(* Logix 5000 project; controller TFF vendor 1 type 14 code 107 rev 34.11; software revision 34.03; part 35 of 36 *)
(* tags used below, declared in another part *)
   Config : Configuration;   // Index Array used in configuration routines
   Index : DINT;   // Index
   FirstScanComplete : BOOL;   // First Scan Complete Flag
   FlowPath : FlowPath[64];   // Flow Path Array
   FlowPathControl : FlowPathControl;   // Flow Path Control
   FlowPathSetup : FlowPathSetup;   // Flow Path Setup Data
   LI001 : ALIAS FOR AnalogPoint[44];   // Feed Bag Volume
   LI001Alarm : ALIAS FOR AlarmAnalog[44];   // Feed Bag Volume Alarm
   Phase0 : ALIAS FOR Phase[0];   // Phase 0
   SysControl : SysControl;   // General system status and command
   Tank : TankManagement;   // Tank Management
   Valve : Valve[100];   // Valve Array
   ValveControl : ValveControl;   // Valve Control
   WI001 : ALIAS FOR AnalogPoint[15];   // Feed Bag Weight
   WI001Alarm : ALIAS FOR AlarmAnalog[15];   // Feed Bag Weight Alarm
(* Process, continued *)

ROUTINE TankRange   (* ladder *)
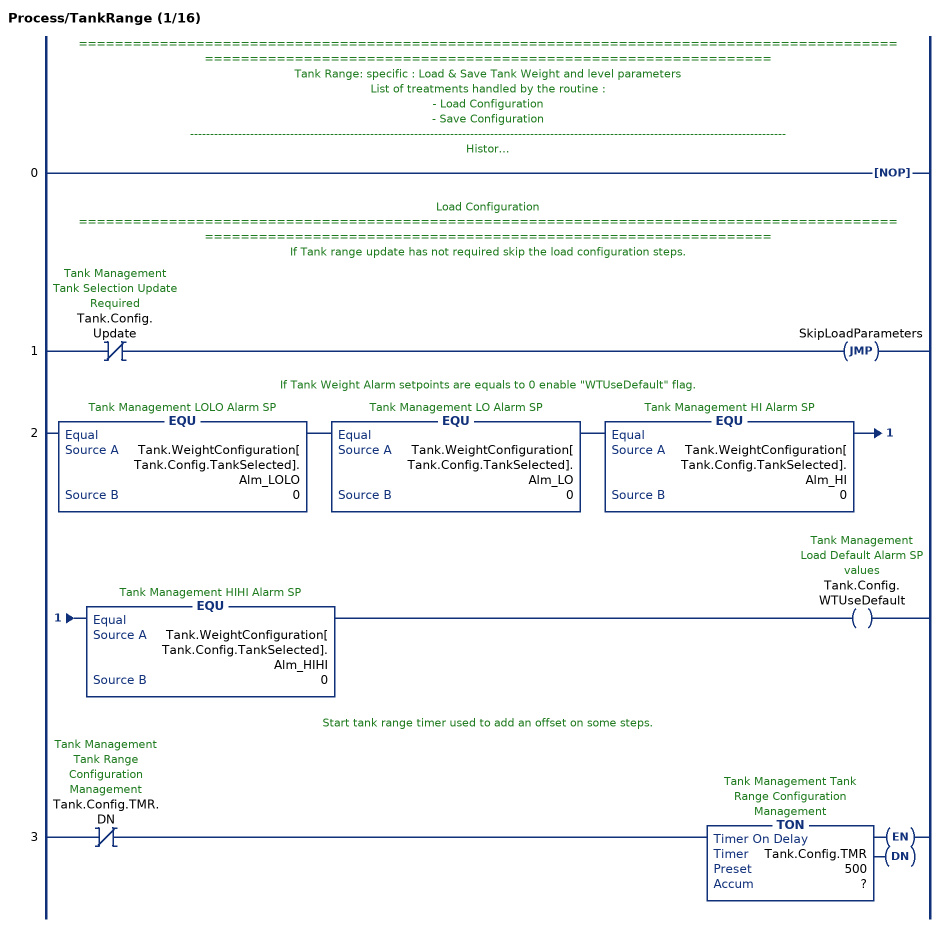
   // ==========================================================================================================================================================
   //                                                                                                                                 Tank Range: specific : Load & Save Tank Weight and level parameters
   //                                                     List of treatments handled by the routine :
   //                                                          - Load Configuration
   //                                                          - Save Configuration
   //                                                     -----------------------------------------------------------------------------------------------------------------------------------------------------
   //                                                     History
   //                                                          2019-AUG-13 - Actemium - B. Roch - Initial version for Candidate Release 3.00.00.00.a
   // ==========================================================================================================================================================
   0: NOP();
   // Load Configuration
   // ==========================================================================================================================================================
   // If Tank range update has not required skip the load configuration steps.
   1: XIO(Tank.Config.Update)JMP(SkipLoadParameters);
   // If Tank Weight Alarm setpoints are equals to 0 enable "WTUseDefault" flag.
   2: EQU(Tank.WeightConfiguration[Tank.Config.TankSelected].Alm_LOLO,0)EQU(Tank.WeightConfiguration[Tank.Config.TankSelected].Alm_LO,0)EQU(Tank.WeightConfiguration[Tank.Config.TankSelected].Alm_HI,0)EQU(Tank.WeightConfiguration[Tank.Config.TankSelected].Alm_HIHI,0)OTE(Tank.Config.WTUseDefault);
   // Start tank range timer used to add an offset on some steps.
   3: XIO(Tank.Config.TMR.DN)TON(Tank.Config.TMR,?,?);
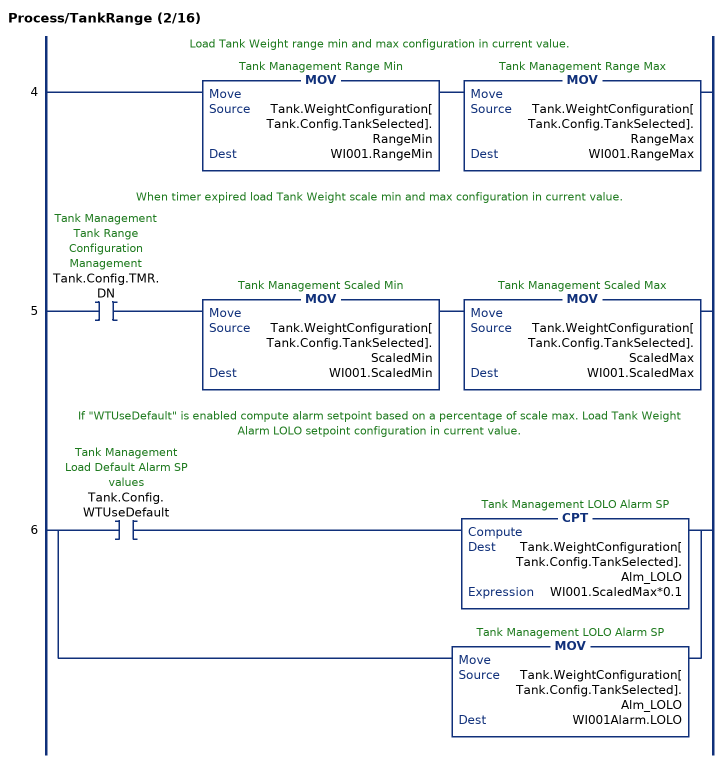
   // Load Tank Weight range min and max configuration in current value.
   4: MOV(Tank.WeightConfiguration[Tank.Config.TankSelected].RangeMin,WI001.RangeMin)MOV(Tank.WeightConfiguration[Tank.Config.TankSelected].RangeMax,WI001.RangeMax);
   // When timer expired load Tank Weight scale min and max configuration in current value.
   5: XIC(Tank.Config.TMR.DN)MOV(Tank.WeightConfiguration[Tank.Config.TankSelected].ScaledMin,WI001.ScaledMin)MOV(Tank.WeightConfiguration[Tank.Config.TankSelected].ScaledMax,WI001.ScaledMax);
   // If "WTUseDefault" is enabled compute alarm setpoint based on a percentage of scale max. Load Tank Weight Alarm LOLO setpoint configuration in current value.
   6: [XIC(Tank.Config.WTUseDefault) CPT(Tank.WeightConfiguration[Tank.Config.TankSelected].Alm_LOLO,WI001.ScaledMax*0.1) ,MOV(Tank.WeightConfiguration[Tank.Config.TankSelected].Alm_LOLO,WI001Alarm.LOLO) ];
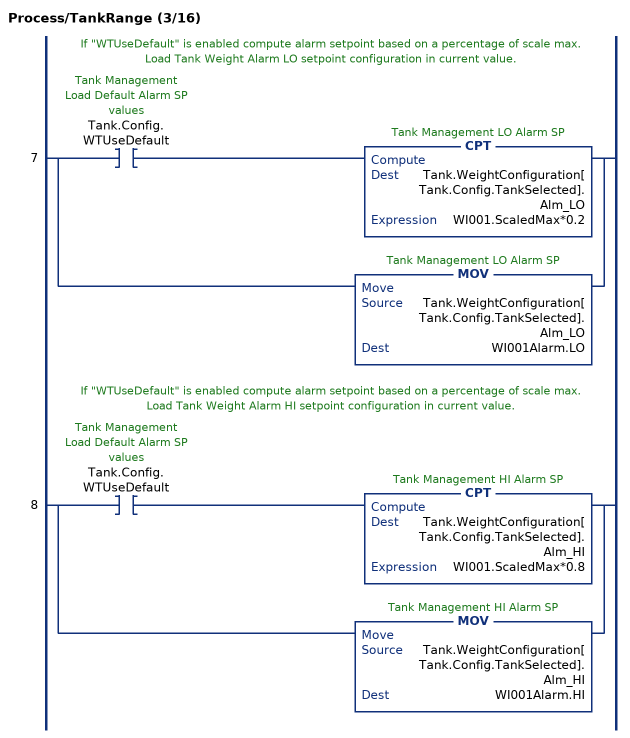
   // If "WTUseDefault" is enabled compute alarm setpoint based on a percentage of scale max. Load Tank Weight Alarm LO setpoint configuration in current value.
   7: [XIC(Tank.Config.WTUseDefault) CPT(Tank.WeightConfiguration[Tank.Config.TankSelected].Alm_LO,WI001.ScaledMax*0.2) ,MOV(Tank.WeightConfiguration[Tank.Config.TankSelected].Alm_LO,WI001Alarm.LO) ];
   // If "WTUseDefault" is enabled compute alarm setpoint based on a percentage of scale max. Load Tank Weight Alarm HI setpoint configuration in current value.
   8: [XIC(Tank.Config.WTUseDefault) CPT(Tank.WeightConfiguration[Tank.Config.TankSelected].Alm_HI,WI001.ScaledMax*0.8) ,MOV(Tank.WeightConfiguration[Tank.Config.TankSelected].Alm_HI,WI001Alarm.HI) ];
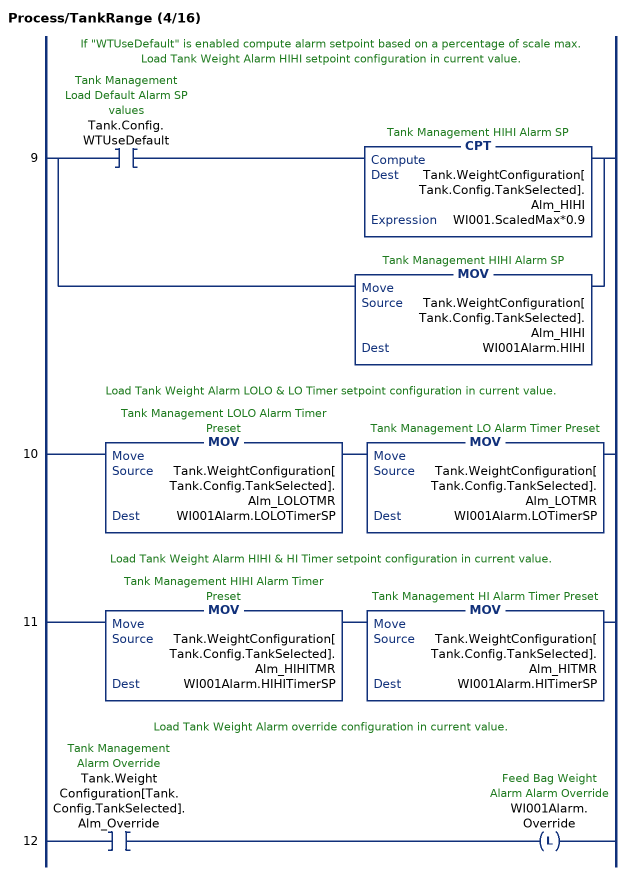
   // If "WTUseDefault" is enabled compute alarm setpoint based on a percentage of scale max. Load Tank Weight Alarm HIHI setpoint configuration in current value.
   9: [XIC(Tank.Config.WTUseDefault) CPT(Tank.WeightConfiguration[Tank.Config.TankSelected].Alm_HIHI,WI001.ScaledMax*0.9) ,MOV(Tank.WeightConfiguration[Tank.Config.TankSelected].Alm_HIHI,WI001Alarm.HIHI) ];
   // Load Tank Weight Alarm LOLO & LO Timer setpoint configuration in current value.
   10: MOV(Tank.WeightConfiguration[Tank.Config.TankSelected].Alm_LOLOTMR,WI001Alarm.LOLOTimerSP)MOV(Tank.WeightConfiguration[Tank.Config.TankSelected].Alm_LOTMR,WI001Alarm.LOTimerSP);
   // Load Tank Weight Alarm HIHI & HI Timer setpoint configuration in current value.
   11: MOV(Tank.WeightConfiguration[Tank.Config.TankSelected].Alm_HIHITMR,WI001Alarm.HIHITimerSP)MOV(Tank.WeightConfiguration[Tank.Config.TankSelected].Alm_HITMR,WI001Alarm.HITimerSP);
   // Load Tank Weight Alarm override configuration in current value.
   12: XIC(Tank.WeightConfiguration[Tank.Config.TankSelected].Alm_Override)OTL(WI001Alarm.Override);
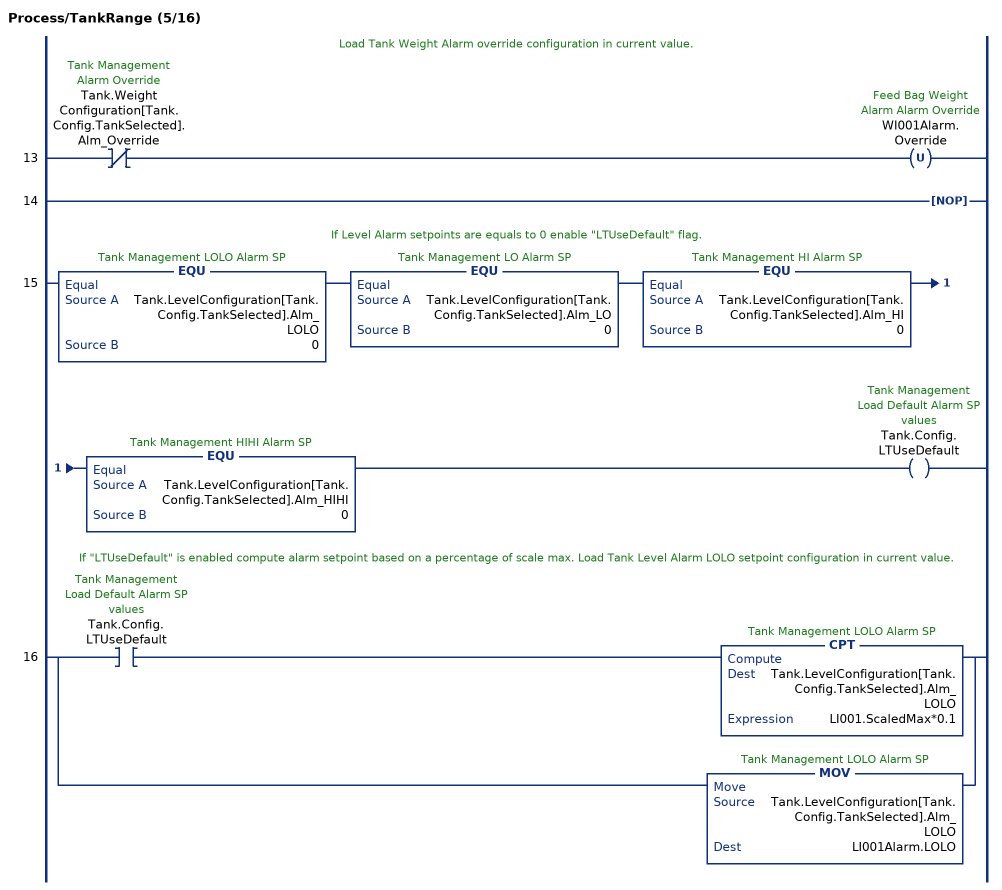
   // Load Tank Weight Alarm override configuration in current value.
   13: XIO(Tank.WeightConfiguration[Tank.Config.TankSelected].Alm_Override)OTU(WI001Alarm.Override);
   14: NOP();
   // If Level Alarm setpoints are equals to 0 enable "LTUseDefault" flag.
   15: EQU(Tank.LevelConfiguration[Tank.Config.TankSelected].Alm_LOLO,0)EQU(Tank.LevelConfiguration[Tank.Config.TankSelected].Alm_LO,0)EQU(Tank.LevelConfiguration[Tank.Config.TankSelected].Alm_HI,0)EQU(Tank.LevelConfiguration[Tank.Config.TankSelected].Alm_HIHI,0)OTE(Tank.Config.LTUseDefault);
   // If "LTUseDefault" is enabled compute alarm setpoint based on a percentage of scale max. Load Tank Level Alarm LOLO setpoint configuration in current value.
   16: [XIC(Tank.Config.LTUseDefault) CPT(Tank.LevelConfiguration[Tank.Config.TankSelected].Alm_LOLO,LI001.ScaledMax*0.1) ,MOV(Tank.LevelConfiguration[Tank.Config.TankSelected].Alm_LOLO,LI001Alarm.LOLO) ];
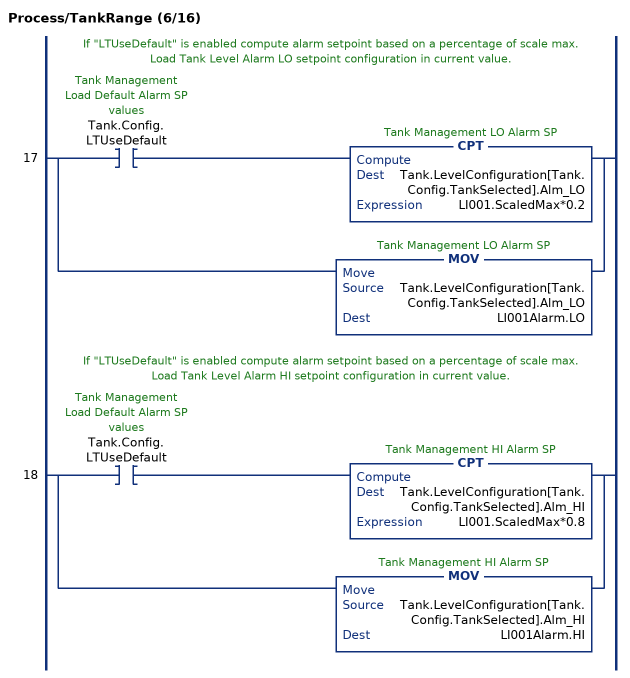
   // If "LTUseDefault" is enabled compute alarm setpoint based on a percentage of scale max. Load Tank Level Alarm LO setpoint configuration in current value.
   17: [XIC(Tank.Config.LTUseDefault) CPT(Tank.LevelConfiguration[Tank.Config.TankSelected].Alm_LO,LI001.ScaledMax*0.2) ,MOV(Tank.LevelConfiguration[Tank.Config.TankSelected].Alm_LO,LI001Alarm.LO) ];
   // If "LTUseDefault" is enabled compute alarm setpoint based on a percentage of scale max. Load Tank Level Alarm HI setpoint configuration in current value.
   18: [XIC(Tank.Config.LTUseDefault) CPT(Tank.LevelConfiguration[Tank.Config.TankSelected].Alm_HI,LI001.ScaledMax*0.8) ,MOV(Tank.LevelConfiguration[Tank.Config.TankSelected].Alm_HI,LI001Alarm.HI) ];
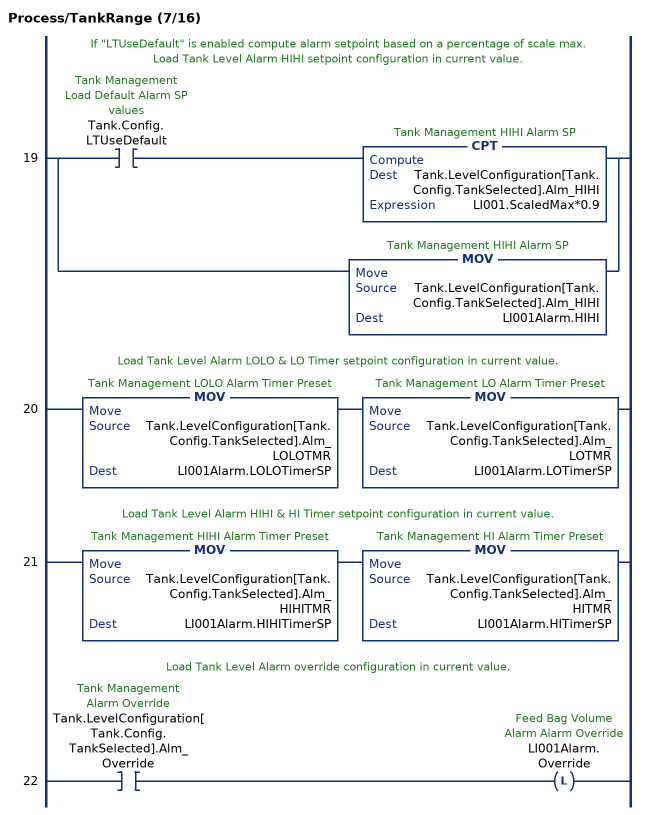
   // If "LTUseDefault" is enabled compute alarm setpoint based on a percentage of scale max. Load Tank Level Alarm HIHI setpoint configuration in current value.
   19: [XIC(Tank.Config.LTUseDefault) CPT(Tank.LevelConfiguration[Tank.Config.TankSelected].Alm_HIHI,LI001.ScaledMax*0.9) ,MOV(Tank.LevelConfiguration[Tank.Config.TankSelected].Alm_HIHI,LI001Alarm.HIHI) ];
   // Load Tank Level Alarm LOLO & LO Timer setpoint configuration in current value.
   20: MOV(Tank.LevelConfiguration[Tank.Config.TankSelected].Alm_LOLOTMR,LI001Alarm.LOLOTimerSP)MOV(Tank.LevelConfiguration[Tank.Config.TankSelected].Alm_LOTMR,LI001Alarm.LOTimerSP);
   // Load Tank Level Alarm HIHI & HI Timer setpoint configuration in current value.
   21: MOV(Tank.LevelConfiguration[Tank.Config.TankSelected].Alm_HIHITMR,LI001Alarm.HIHITimerSP)MOV(Tank.LevelConfiguration[Tank.Config.TankSelected].Alm_HITMR,LI001Alarm.HITimerSP);
   // Load Tank Level Alarm override configuration in current value.
   22: XIC(Tank.LevelConfiguration[Tank.Config.TankSelected].Alm_Override)OTL(LI001Alarm.Override);
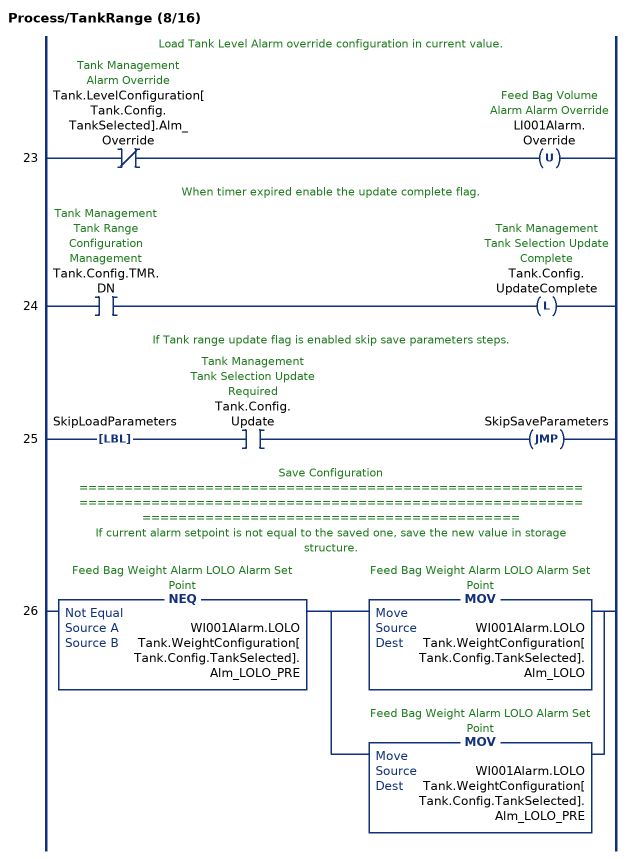
   // Load Tank Level Alarm override configuration in current value.
   23: XIO(Tank.LevelConfiguration[Tank.Config.TankSelected].Alm_Override)OTU(LI001Alarm.Override);
   // When timer expired enable the update complete flag.
   24: XIC(Tank.Config.TMR.DN)OTL(Tank.Config.UpdateComplete);
   // If Tank range update flag is enabled skip save parameters steps.
   25: LBL(SkipLoadParameters)XIC(Tank.Config.Update)JMP(SkipSaveParameters);
   // Save Configuration
   // ==========================================================================================================================================================
   // If current alarm setpoint is not equal to the saved one, save the new value in storage structure.
   26: NEQ(WI001Alarm.LOLO,Tank.WeightConfiguration[Tank.Config.TankSelected].Alm_LOLO_PRE)[MOV(WI001Alarm.LOLO,Tank.WeightConfiguration[Tank.Config.TankSelected].Alm_LOLO) ,MOV(WI001Alarm.LOLO,Tank.WeightConfiguration[Tank.Config.TankSelected].Alm_LOLO_PRE) ];
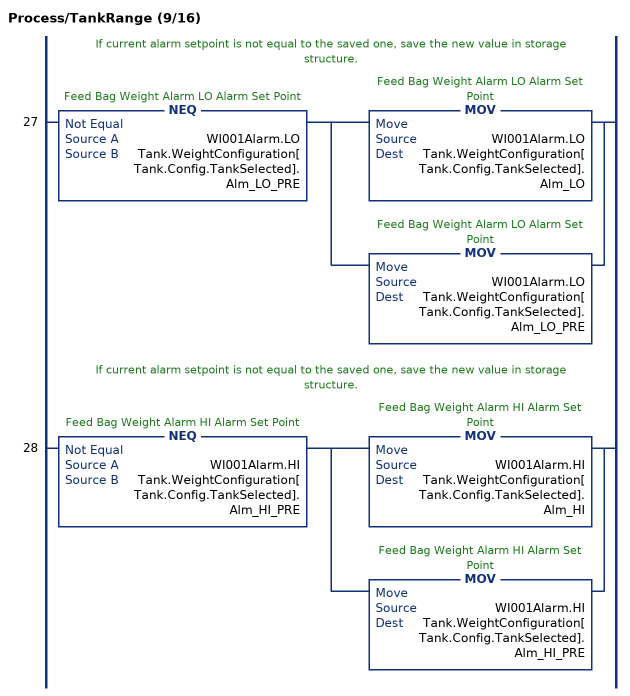
   // If current alarm setpoint is not equal to the saved one, save the new value in storage structure.
   27: NEQ(WI001Alarm.LO,Tank.WeightConfiguration[Tank.Config.TankSelected].Alm_LO_PRE)[MOV(WI001Alarm.LO,Tank.WeightConfiguration[Tank.Config.TankSelected].Alm_LO) ,MOV(WI001Alarm.LO,Tank.WeightConfiguration[Tank.Config.TankSelected].Alm_LO_PRE) ];
   // If current alarm setpoint is not equal to the saved one, save the new value in storage structure.
   28: NEQ(WI001Alarm.HI,Tank.WeightConfiguration[Tank.Config.TankSelected].Alm_HI_PRE)[MOV(WI001Alarm.HI,Tank.WeightConfiguration[Tank.Config.TankSelected].Alm_HI) ,MOV(WI001Alarm.HI,Tank.WeightConfiguration[Tank.Config.TankSelected].Alm_HI_PRE) ];
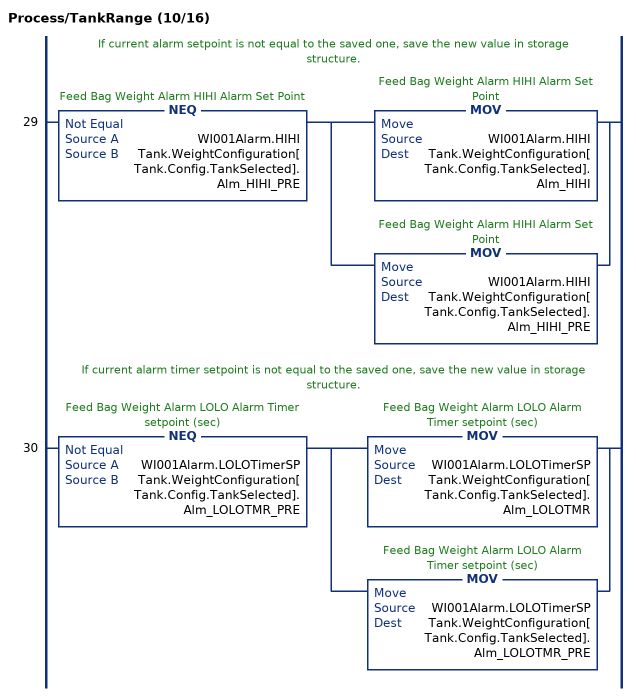
   // If current alarm setpoint is not equal to the saved one, save the new value in storage structure.
   29: NEQ(WI001Alarm.HIHI,Tank.WeightConfiguration[Tank.Config.TankSelected].Alm_HIHI_PRE)[MOV(WI001Alarm.HIHI,Tank.WeightConfiguration[Tank.Config.TankSelected].Alm_HIHI) ,MOV(WI001Alarm.HIHI,Tank.WeightConfiguration[Tank.Config.TankSelected].Alm_HIHI_PRE) ];
   // If current alarm timer setpoint is not equal to the saved one, save the new value in storage structure.
   30: NEQ(WI001Alarm.LOLOTimerSP,Tank.WeightConfiguration[Tank.Config.TankSelected].Alm_LOLOTMR_PRE)[MOV(WI001Alarm.LOLOTimerSP,Tank.WeightConfiguration[Tank.Config.TankSelected].Alm_LOLOTMR) ,MOV(WI001Alarm.LOLOTimerSP,Tank.WeightConfiguration[Tank.Config.TankSelected].Alm_LOLOTMR_PRE) ];
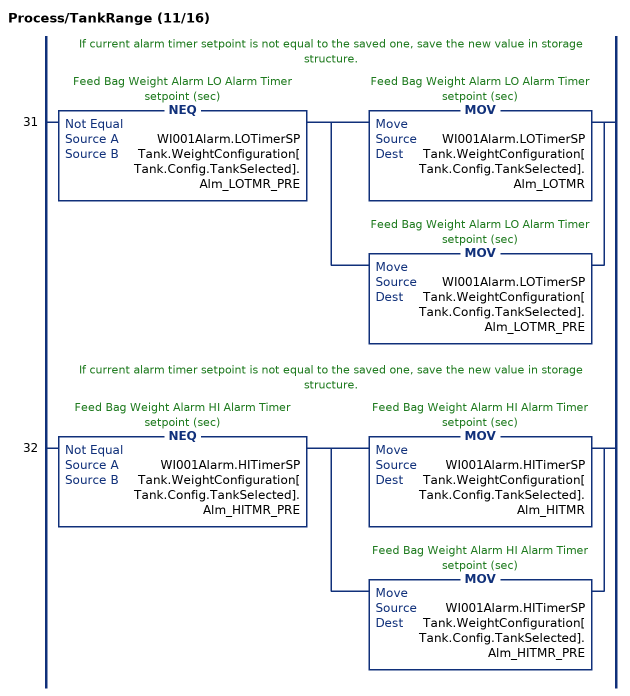
   // If current alarm timer setpoint is not equal to the saved one, save the new value in storage structure.
   31: NEQ(WI001Alarm.LOTimerSP,Tank.WeightConfiguration[Tank.Config.TankSelected].Alm_LOTMR_PRE)[MOV(WI001Alarm.LOTimerSP,Tank.WeightConfiguration[Tank.Config.TankSelected].Alm_LOTMR) ,MOV(WI001Alarm.LOTimerSP,Tank.WeightConfiguration[Tank.Config.TankSelected].Alm_LOTMR_PRE) ];
   // If current alarm timer setpoint is not equal to the saved one, save the new value in storage structure.
   32: NEQ(WI001Alarm.HITimerSP,Tank.WeightConfiguration[Tank.Config.TankSelected].Alm_HITMR_PRE)[MOV(WI001Alarm.HITimerSP,Tank.WeightConfiguration[Tank.Config.TankSelected].Alm_HITMR) ,MOV(WI001Alarm.HITimerSP,Tank.WeightConfiguration[Tank.Config.TankSelected].Alm_HITMR_PRE) ];
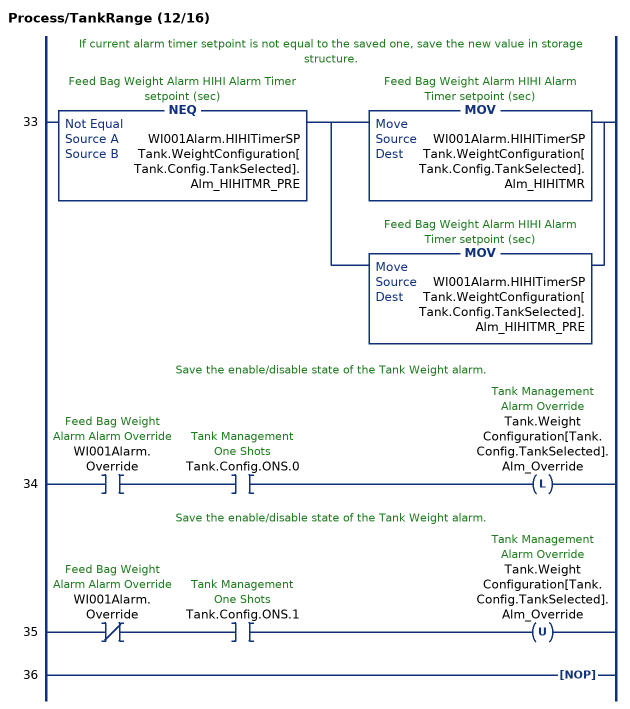
   // If current alarm timer setpoint is not equal to the saved one, save the new value in storage structure.
   33: NEQ(WI001Alarm.HIHITimerSP,Tank.WeightConfiguration[Tank.Config.TankSelected].Alm_HIHITMR_PRE)[MOV(WI001Alarm.HIHITimerSP,Tank.WeightConfiguration[Tank.Config.TankSelected].Alm_HIHITMR) ,MOV(WI001Alarm.HIHITimerSP,Tank.WeightConfiguration[Tank.Config.TankSelected].Alm_HIHITMR_PRE) ];
   // Save the enable/disable state of the Tank Weight alarm.
   34: XIC(WI001Alarm.Override)XIC(Tank.Config.ONS.0)OTL(Tank.WeightConfiguration[Tank.Config.TankSelected].Alm_Override);
   // Save the enable/disable state of the Tank Weight alarm.
   35: XIO(WI001Alarm.Override)XIC(Tank.Config.ONS.1)OTU(Tank.WeightConfiguration[Tank.Config.TankSelected].Alm_Override);
   36: NOP();
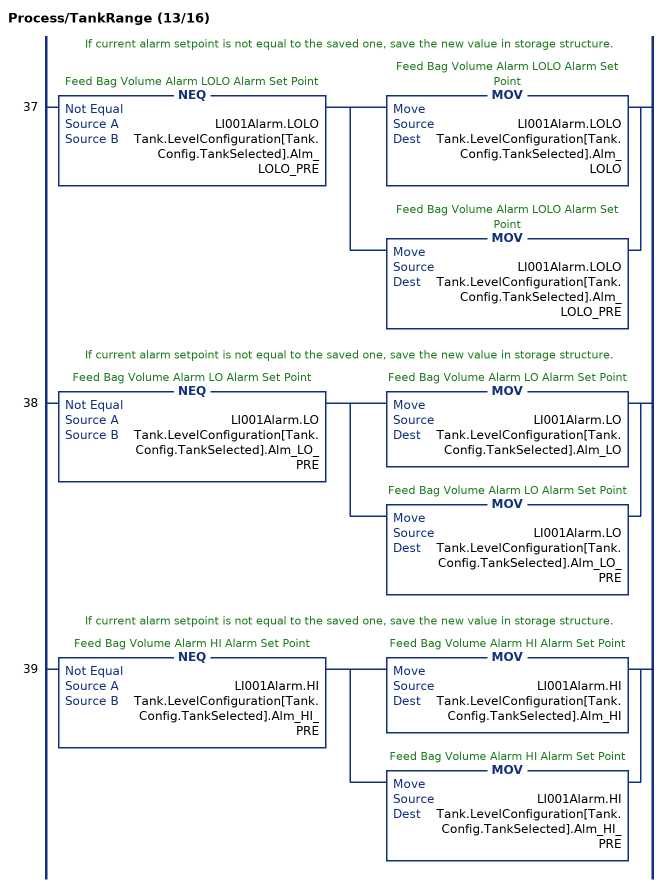
   // If current alarm setpoint is not equal to the saved one, save the new value in storage structure.
   37: NEQ(LI001Alarm.LOLO,Tank.LevelConfiguration[Tank.Config.TankSelected].Alm_LOLO_PRE)[MOV(LI001Alarm.LOLO,Tank.LevelConfiguration[Tank.Config.TankSelected].Alm_LOLO) ,MOV(LI001Alarm.LOLO,Tank.LevelConfiguration[Tank.Config.TankSelected].Alm_LOLO_PRE) ];
   // If current alarm setpoint is not equal to the saved one, save the new value in storage structure.
   38: NEQ(LI001Alarm.LO,Tank.LevelConfiguration[Tank.Config.TankSelected].Alm_LO_PRE)[MOV(LI001Alarm.LO,Tank.LevelConfiguration[Tank.Config.TankSelected].Alm_LO) ,MOV(LI001Alarm.LO,Tank.LevelConfiguration[Tank.Config.TankSelected].Alm_LO_PRE) ];
   // If current alarm setpoint is not equal to the saved one, save the new value in storage structure.
   39: NEQ(LI001Alarm.HI,Tank.LevelConfiguration[Tank.Config.TankSelected].Alm_HI_PRE)[MOV(LI001Alarm.HI,Tank.LevelConfiguration[Tank.Config.TankSelected].Alm_HI) ,MOV(LI001Alarm.HI,Tank.LevelConfiguration[Tank.Config.TankSelected].Alm_HI_PRE) ];
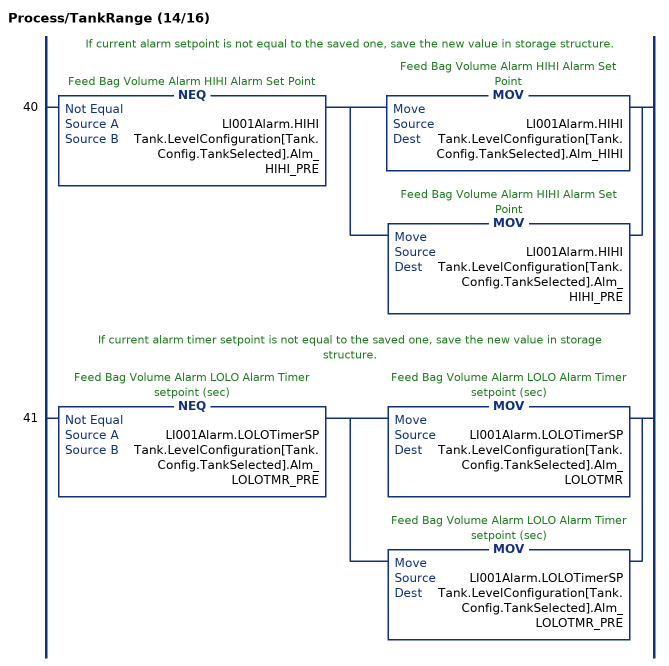
   // If current alarm setpoint is not equal to the saved one, save the new value in storage structure.
   40: NEQ(LI001Alarm.HIHI,Tank.LevelConfiguration[Tank.Config.TankSelected].Alm_HIHI_PRE)[MOV(LI001Alarm.HIHI,Tank.LevelConfiguration[Tank.Config.TankSelected].Alm_HIHI) ,MOV(LI001Alarm.HIHI,Tank.LevelConfiguration[Tank.Config.TankSelected].Alm_HIHI_PRE) ];
   // If current alarm timer setpoint is not equal to the saved one, save the new value in storage structure.
   41: NEQ(LI001Alarm.LOLOTimerSP,Tank.LevelConfiguration[Tank.Config.TankSelected].Alm_LOLOTMR_PRE)[MOV(LI001Alarm.LOLOTimerSP,Tank.LevelConfiguration[Tank.Config.TankSelected].Alm_LOLOTMR) ,MOV(LI001Alarm.LOLOTimerSP,Tank.LevelConfiguration[Tank.Config.TankSelected].Alm_LOLOTMR_PRE) ];
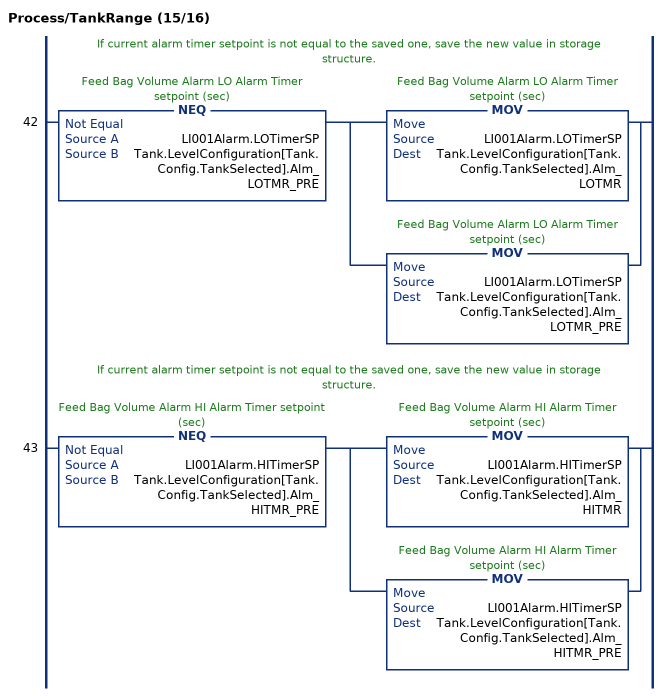
   // If current alarm timer setpoint is not equal to the saved one, save the new value in storage structure.
   42: NEQ(LI001Alarm.LOTimerSP,Tank.LevelConfiguration[Tank.Config.TankSelected].Alm_LOTMR_PRE)[MOV(LI001Alarm.LOTimerSP,Tank.LevelConfiguration[Tank.Config.TankSelected].Alm_LOTMR) ,MOV(LI001Alarm.LOTimerSP,Tank.LevelConfiguration[Tank.Config.TankSelected].Alm_LOTMR_PRE) ];
   // If current alarm timer setpoint is not equal to the saved one, save the new value in storage structure.
   43: NEQ(LI001Alarm.HITimerSP,Tank.LevelConfiguration[Tank.Config.TankSelected].Alm_HITMR_PRE)[MOV(LI001Alarm.HITimerSP,Tank.LevelConfiguration[Tank.Config.TankSelected].Alm_HITMR) ,MOV(LI001Alarm.HITimerSP,Tank.LevelConfiguration[Tank.Config.TankSelected].Alm_HITMR_PRE) ];
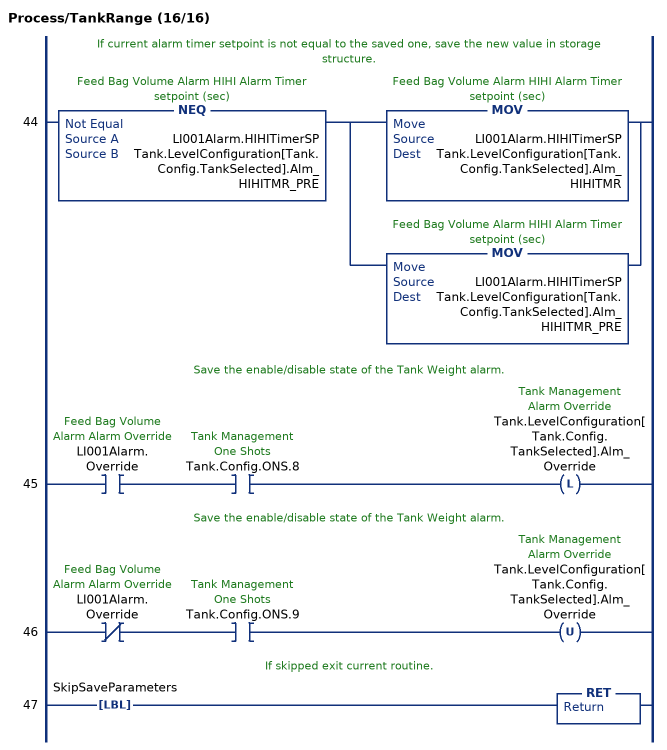
   // If current alarm timer setpoint is not equal to the saved one, save the new value in storage structure.
   44: NEQ(LI001Alarm.HIHITimerSP,Tank.LevelConfiguration[Tank.Config.TankSelected].Alm_HIHITMR_PRE)[MOV(LI001Alarm.HIHITimerSP,Tank.LevelConfiguration[Tank.Config.TankSelected].Alm_HIHITMR) ,MOV(LI001Alarm.HIHITimerSP,Tank.LevelConfiguration[Tank.Config.TankSelected].Alm_HIHITMR_PRE) ];
   // Save the enable/disable state of the Tank Weight alarm.
   45: XIC(LI001Alarm.Override)XIC(Tank.Config.ONS.8)OTL(Tank.LevelConfiguration[Tank.Config.TankSelected].Alm_Override);
   // Save the enable/disable state of the Tank Weight alarm.
   46: XIO(LI001Alarm.Override)XIC(Tank.Config.ONS.9)OTU(Tank.LevelConfiguration[Tank.Config.TankSelected].Alm_Override);
   // If skipped exit current routine.
   47: LBL(SkipSaveParameters)RET();
END_ROUTINE

ROUTINE Valve   (* ladder *)
// Valve Control Routine
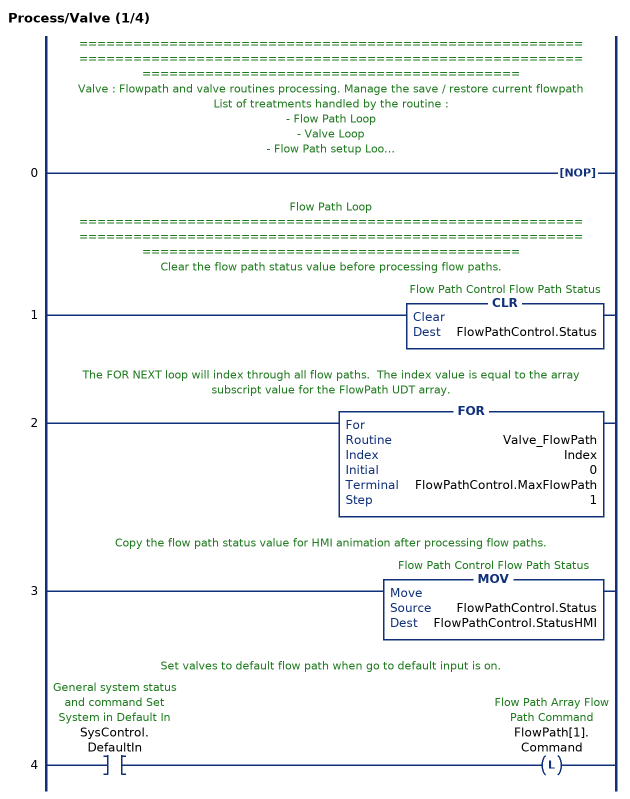
   // ==========================================================================================================================================================
   //                                                                                    Valve : Flowpath and valve routines processing. Manage the save / restore current flowpath
   //                                                     List of treatments handled by the routine :
   //                                                          - Flow Path Loop
   //                                                          - Valve Loop
   //                                                          - Flow Path setup Loop
   //                                                          - Save/restore current flowpath
   //                                                     -----------------------------------------------------------------------------------------------------------------------------------------------------
   //                                                     History
   //                                                          2019-AUG-13 - Actemium - B. Roch - Initial version for Candidate Release 3.00.00.00.a
   // 		2023-FEB-09 - DAVIDSON - Ch. ARBOGAST - Modification for Candidate Release 2.02.00.00.b
   //                                                - Rung 10 to 13; change save flowpath logic, making it resilient from power failure when in hold.
   // =============================================================================================================
   0: NOP();
   // Flow Path Loop
   // ==========================================================================================================================================================
   // Clear the flow path status value before processing flow paths.
   1: CLR(FlowPathControl.Status);
   // The FOR NEXT loop will index through all flow paths.  The index value is equal to the array subscript value for the FlowPath UDT array.
   2: FOR(Valve_FlowPath,Index,0,FlowPathControl.MaxFlowPath,1);
   // Copy the flow path status value for HMI animation after processing flow paths.
   3: MOV(FlowPathControl.Status,FlowPathControl.StatusHMI);
   // Set valves to default flow path when go to default input is on.
   4: XIC(SysControl.DefaultIn)OTL(FlowPath[1].Command);
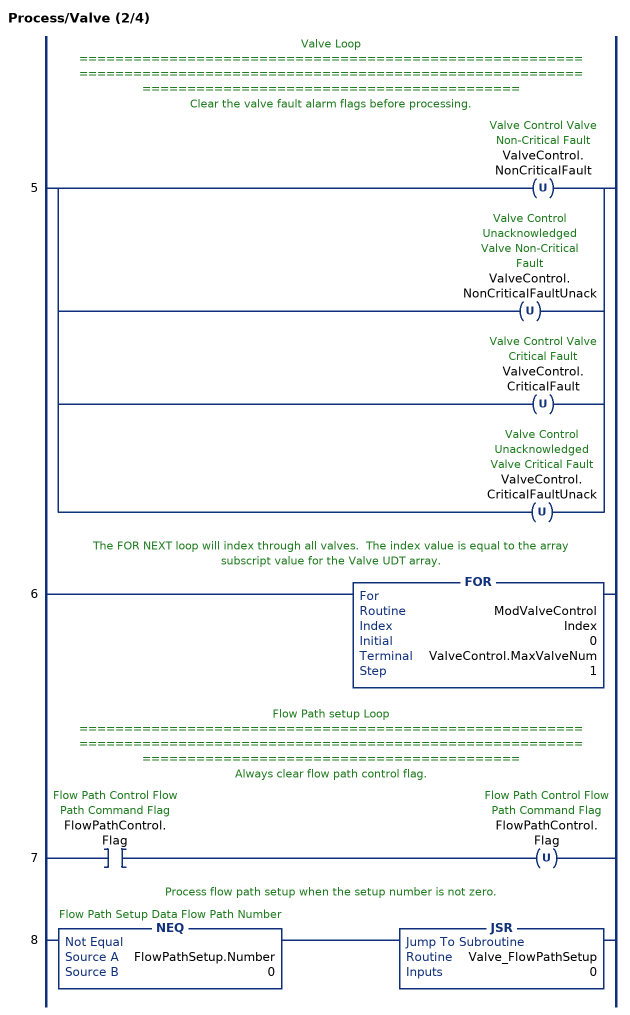
   // Valve Loop
   // ==========================================================================================================================================================
   // Clear the valve fault alarm flags before processing.
   5: [OTU(ValveControl.NonCriticalFault) ,OTU(ValveControl.NonCriticalFaultUnack) ,OTU(ValveControl.CriticalFault) ,OTU(ValveControl.CriticalFaultUnack) ];
   // The FOR NEXT loop will index through all valves.  The index value is equal to the array subscript value for the Valve UDT array.
   6: FOR(ModValveControl,Index,0,ValveControl.MaxValveNum,1);
   // Flow Path setup Loop
   // ==========================================================================================================================================================
   // Always clear flow path control flag.
   7: XIC(FlowPathControl.Flag)OTU(FlowPathControl.Flag);
   // Process flow path setup when the setup number is not zero.
   8: NEQ(FlowPathSetup.Number,0)JSR(Valve_FlowPathSetup,0);
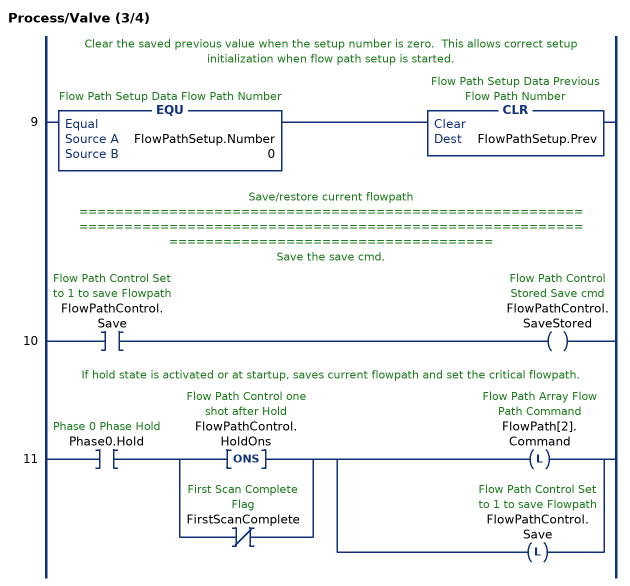
   // Clear the saved previous value when the setup number is zero.  This allows correct setup initialization when flow path setup is started.
   9: EQU(FlowPathSetup.Number,0)CLR(FlowPathSetup.Prev);
   // Save/restore current flowpath
   // ====================================================================================================================================================
   // Save the save cmd.
   10: XIC(FlowPathControl.Save)OTE(FlowPathControl.SaveStored);
   // If hold state is activated or at startup, saves current flowpath and set the critical flowpath.
   11: XIC(Phase0.Hold)[ONS(FlowPathControl.HoldOns) ,XIO(FirstScanComplete) ][OTL(FlowPath[2].Command) ,OTL(FlowPathControl.Save) ];
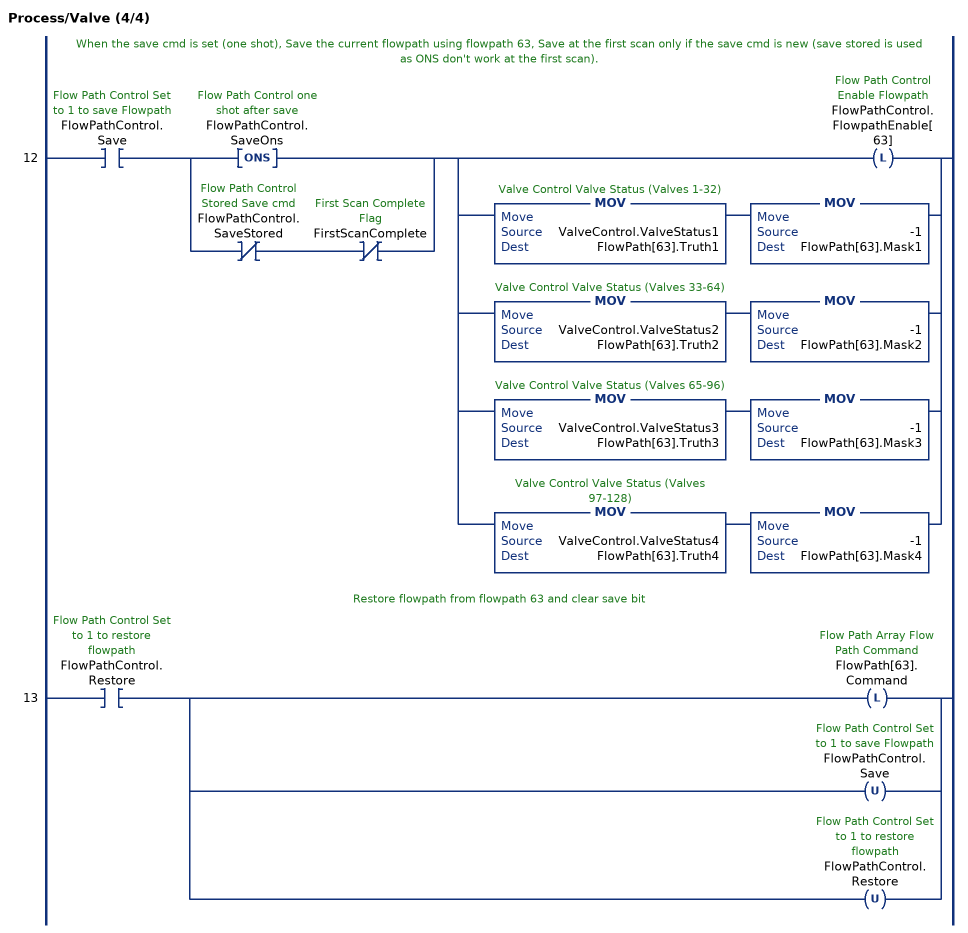
   // When the save cmd is set (one shot), Save the current flowpath using flowpath 63, Save at the first scan only if the save cmd is new (save stored is used as ONS don't work at the first scan).
   12: XIC(FlowPathControl.Save)[ONS(FlowPathControl.SaveOns) ,XIO(FlowPathControl.SaveStored) XIO(FirstScanComplete) ][OTL(FlowPathControl.FlowpathEnable[63]) ,MOV(ValveControl.ValveStatus1,FlowPath[63].Truth1) MOV(-1,FlowPath[63].Mask1) ,MOV(ValveControl.ValveStatus2,FlowPath[63].Truth2) MOV(-1,FlowPath[63].Mask2) ,MOV(ValveControl.ValveStatus3,FlowPath[63].Truth3) MOV(-1,FlowPath[63].Mask3) ,MOV(ValveControl.ValveStatus4,FlowPath[63].Truth4) MOV(-1,FlowPath[63].Mask4) ];
   // Restore flowpath from flowpath 63 and clear save bit
   13: XIC(FlowPathControl.Restore)[OTL(FlowPath[63].Command) ,OTU(FlowPathControl.Save) ,OTU(FlowPathControl.Restore) ];
END_ROUTINE
